TYPE ST_AnalogSensor_Diag :
STRUCT
	NoOfSamples : USINT;
	error		: BIT;
	underrange	: BIT;
	overrange	: BIT;
	diag		: BIT;
	limit1		: BIT;
	limit2		: BIT;

END_STRUCT
END_TYPE

(* stored: Version 1.1.0.1
   DUT ST_AnalogSensor_Diag: Id {3c6fafaa-246d-4953-899c-63b110adeddb} *)
